Fanuc KAREL source: KO00015.KL

PROGRAM KO00015
%NOLOCKGROUP
VAR
  P1: XYZWPR
  P2: XYZWPR
  P3: XYZWPR
  P4: XYZWPR
  OUT: XYZWPREXT
BEGIN
  OUT = FRAME(P1, P2, P3, P4)
END KO00015
